KUKA KRL program: SpeedProg.src

&ACCESS RVP
&REL 1
&PARAM TEMPLATE = C:\KRC\Roboter\Template\vorgabe
&PARAM EDITMASK = *
DEF SpeedProg ( )


; GLOBAL INTERRUPT DECL 3 WHEN $STOPMESS==TRUE DO IR_STOPM ( )
; INTERRUPT ON 3

;FOLD Initialise and set default speed
BAS (#INITMOV,0)
BAS (#VEL_PTP,100)
BAS (#ACC_PTP,20)
$VEL.CP=0.2
BAS (#TOOL,0)
BAS (#BASE,0)
;ENDFOLD

;;FOLD STARTPOS
;$BWDSTART = FALSE
;PDAT_ACT = PDEFAULT
;BAS(#PTP_DAT)
;FDAT_ACT = {TOOL_NO 0,BASE_NO 0,IPO_FRAME #BASE}
;BAS(#FRAMES)
;;ENDFOLD

$ADVANCE = 5

;FOLD ---- Quickly skip BCO ----
; PTP $AXIS_ACT
;ENDFOLD

;FOLD ---- GO HOME ----
; PTP {A1 0.000, A2 -90.000, A3 90.000, A4 0.000, A5 0.000, A6 0.000, E1 0, E2 0, E3 0, E4 0, E5 0, E6 0}
;ENDFOLD


; Program generated by RoboDK v6.0.7 for KUKA KR 6 R700 Z200 on XX/XX/XXXX 18:00:00
; Using nominal kinematics.
; ---- Setting reference (Base) ----
$BASE = {FRAME: X 1234.570,Y -98.765,Z 50.500,A 30.000,B 0.000,C 0.000}
; --------------------------
; ---- Setting tool (TCP) ----
$TOOL = {FRAME: X 10.000,Y 20.000,Z 150.000,A 0.000,B 0.000,C 0.000}
; --------------------------
$APO.CPTP = 0
$APO.CDIS = 0.300
$VEL.CP = 0.00100
LIN {X -607.850,Y 543.849,Z 363.215,A 150.000,B 50.000,C -165.000} C_DIS
$VEL.ORI1 = 1.00000
$VEL.ORI2 = 1.00000
PTP {A1 10.00000,A2 -20.00000,A3 50.00000,A4 0.00000,A5 60.00000,A6 30.00000} C_PTP
$APO.CPTP = 1
$APO.CDIS = 1.000
$VEL.CP = 0.01230
LIN {X -640.584,Y 506.980,Z 371.534,A 150.000,B 50.000,C -165.000} C_DIS
$VEL.ORI1 = 5.50000
$VEL.ORI2 = 5.50000
PTP {A1 30.00000,A2 25.00000,A3 80.00000,A4 0.00000,A5 -15.00000,A6 -45.00000} C_PTP
$APO.CPTP = 2
$APO.CDIS = 2.500
$VEL.CP = 0.09990
LIN {X -607.850,Y 543.849,Z 363.215,A 150.000,B 50.000,C -165.000} C_DIS
$VEL.ORI1 = 20.00000
$VEL.ORI2 = 20.00000
PTP {A1 10.00000,A2 -20.00000,A3 50.00000,A4 0.00000,A5 60.00000,A6 30.00000} C_PTP
$APO.CPTP = 3
$APO.CDIS = 3.700
$VEL.CP = 0.33333
LIN {X -640.584,Y 506.980,Z 371.534,A 150.000,B 50.000,C -165.000} C_DIS
$VEL.ORI1 = 45.00000
$VEL.ORI2 = 45.00000
PTP {A1 30.00000,A2 25.00000,A3 80.00000,A4 0.00000,A5 -15.00000,A6 -45.00000} C_PTP
$APO.CPTP = 6
$APO.CDIS = 6.000
$VEL.CP = 1.00000
LIN {X -607.850,Y 543.849,Z 363.215,A 150.000,B 50.000,C -165.000} C_DIS
$VEL.ORI1 = 90.00000
$VEL.ORI2 = 90.00000
PTP {A1 10.00000,A2 -20.00000,A3 50.00000,A4 0.00000,A5 60.00000,A6 30.00000} C_PTP
$APO.CPTP = 9
$APO.CDIS = 9.000
$VEL.CP = 2.50000
LIN {X -640.584,Y 506.980,Z 371.534,A 150.000,B 50.000,C -165.000} C_DIS
$VEL.ORI1 = 120.00000
$VEL.ORI2 = 120.00000
PTP {A1 30.00000,A2 25.00000,A3 80.00000,A4 0.00000,A5 -15.00000,A6 -45.00000} C_PTP
$APO.CPTP = 15
$APO.CDIS = 15.000
$VEL.CP = 5.00000
LIN {X -607.850,Y 543.849,Z 363.215,A 150.000,B 50.000,C -165.000} C_DIS
$VEL.ORI1 = 180.00000
$VEL.ORI2 = 180.00000
PTP {A1 10.00000,A2 -20.00000,A3 50.00000,A4 0.00000,A5 60.00000,A6 30.00000} C_PTP
$APO.CPTP = 30
$APO.CDIS = 30.000
$VEL.CP = 12.00000
LIN {X -640.584,Y 506.980,Z 371.534,A 150.000,B 50.000,C -165.000} C_DIS
$VEL.ORI1 = 270.00000
$VEL.ORI2 = 270.00000
PTP {A1 30.00000,A2 25.00000,A3 80.00000,A4 0.00000,A5 -15.00000,A6 -45.00000} C_PTP
$APO.CPTP = 75
$APO.CDIS = 75.000
$VEL.CP = 0.00050
LIN {X -607.850,Y 543.849,Z 363.215,A 150.000,B 50.000,C -165.000} C_DIS
$VEL.ORI1 = 400.00000
$VEL.ORI2 = 400.00000
PTP {A1 10.00000,A2 -20.00000,A3 50.00000,A4 0.00000,A5 60.00000,A6 30.00000} C_PTP
$APO.CPTP = 100
$APO.CDIS = 150.000
$VEL.CP = 0.75000
LIN {X -640.584,Y 506.980,Z 371.534,A 150.000,B 50.000,C -165.000} C_DIS
$VEL.ORI1 = 2.25000
$VEL.ORI2 = 2.25000
PTP {A1 30.00000,A2 25.00000,A3 80.00000,A4 0.00000,A5 -15.00000,A6 -45.00000} C_PTP
$ACC.CP = 2.00000
$ACC.ORI1 = 500.00000
$ACC.ORI2 = 500.00000
LIN {X -640.584,Y 506.980,Z 371.534,A 150.000,B 50.000,C -165.000} C_DIS
END
